Fanuc KAREL source: kt00337.KL

-- PROVISIONAL review KL for V770-1; original PC SHA256 64d5e5a973fa8f3921e543dedd4f7200b65e95ac6816eb3c4361195f4e46fa72
-- Incomplete behavior may be omitted. Consult companion uncertainty JSON. Do not deploy.
PROGRAM KT00337
%NOLOCKGROUP
VAR
  B1 : BOOLEAN
  B2 : BOOLEAN
  OUT : BOOLEAN
BEGIN
  -- UNRESOLVED_PC offsets 5-12; opcodes 9D,23
  -- UNRESOLVED_PC offsets 17-24; opcodes 9C,23
  -- UNRESOLVED_PC offsets 29-36; opcodes 9D,23
  -- UNRESOLVED_PC offsets 41-48; opcodes 9C,23
  -- UNRESOLVED_PC offsets 53-72; opcodes 21,21,59,23
  -- UNRESOLVED_PC offsets 77-81; opcodes 7F
END KT00337
